// TIA Portal project "CanvasE2E" (V19)

(* hardware
DEVICE "PLC_1"  S7-1500 station
   slot 0: "导轨_0"  Rack  6ES7 590-1***0-0AA0
   slot 1: "PLC_1"  CPU 1511-1 PN  6ES7 511-1AK01-0AB0  V2.5
      slot 3: "CPU 显示_1"  6ES7591-1AA00-0AA0
      slot 32768: "PROFINET 接口_1"  X1
         slot 32769: "端口_1"  X1 P1
         slot 32770: "端口_2"  X1 P2
*)

// ===== PLC "PLC_1"  CPU 1511-1 PN =====

DATA_BLOCK "iFB_CM_CLAMP_CYL_DRV"   // DB1
{ S7_Optimized_Access := 'TRUE' }
VERSION : 0.1
// stored: InstanceOfName FB_CM_CLAMP_CYL_DRV
"FB_CM_CLAMP_CYL_DRV"
BEGIN
END_DATA_BLOCK

DATA_BLOCK "iFB_EM_CLAMP_SEQ"   // DB2
{ S7_Optimized_Access := 'TRUE' }
VERSION : 0.1
// stored: InstanceOfName FB_EM_CLAMP_SEQ
"FB_EM_CLAMP_SEQ"
BEGIN
END_DATA_BLOCK

DATA_BLOCK "iFB_U_ASSEMBLY_UNIT"   // DB3
{ S7_Optimized_Access := 'TRUE' }
VERSION : 0.1
// stored: InstanceOfName FB_U_ASSEMBLY_UNIT
"FB_U_ASSEMBLY_UNIT"
BEGIN
END_DATA_BLOCK

FUNCTION_BLOCK "PumpCtrl"   // FB1, SCL
{ S7_Optimized_Access := 'TRUE' }
   VAR_INPUT
      Start : Bool;
   END_VAR
   VAR_OUTPUT
      RunOut : Bool;
   END_VAR
   VAR
      Running : Bool;
   END_VAR
BEGIN
       // Network 1: Self-holding logic
       IF #Start THEN
           #Running := TRUE;
       END_IF;
       #RunOut := #Running;
END_FUNCTION_BLOCK

FUNCTION_BLOCK "FB_CM_CLAMP_CYL_DRV"   // FB2, SCL
{ S7_Optimized_Access := 'TRUE' }
   VAR_INPUT
      CmdExtend : Bool;
      CmdRetract : Bool;
      Extended : Bool;
      Retracted : Bool;
   END_VAR
   VAR_OUTPUT
      Q_Extend : Bool;
      Q_Retract : Bool;
      Busy : Bool;
      Done : Bool;
      Error : Bool;
   END_VAR
BEGIN
       // single-writer arbitration + feedback exclusivity
       IF #Extended AND #Retracted THEN
           #Error := TRUE;
           #Q_Extend := FALSE;
           #Q_Retract := FALSE;
       ELSE
           #Error := FALSE;
           #Q_Extend := #CmdExtend AND NOT #CmdRetract;
           #Q_Retract := #CmdRetract AND NOT #CmdExtend;
       END_IF;
       #Busy := #Q_Extend OR #Q_Retract;
END_FUNCTION_BLOCK

FUNCTION_BLOCK "FB_EM_CLAMP_SEQ"   // FB3, SCL
{ S7_Optimized_Access := 'TRUE' }
   VAR_INPUT
      Start : Bool;
      Reset : Bool;
      SafetyPermit : Bool;
      Extended : Bool;
      Retracted : Bool;
   END_VAR
   VAR_OUTPUT
      Busy : Bool;
      Done : Bool;
      Error : Bool;
      StepNo : Int;
      Extend : Bool;
      Retract : Bool;
   END_VAR
   VAR
      "Step" : Int := 0;
      FaultLatch : Bool;
      TON_S_EXTEND : TON_TIME;
      TON_S_HOLD : TON_TIME;
      TON_S_RETRACT : TON_TIME;
   END_VAR
BEGIN
       CASE #Step OF
           0: // S_WAIT 绛夊緟鍚姩
               #Busy := FALSE;
               #Done := FALSE;
               IF #Start AND #SafetyPermit THEN
                   #Step := 10;
               END_IF;
           10: // S_EXTEND 浼稿嚭澶圭揣
               #Busy := TRUE;
               #Extend := TRUE;
               #TON_S_EXTEND(IN := NOT #Extended,
                             PT := T#3000ms);
               IF #Extended THEN
                   #Extend := FALSE;
                   #Step := 20;
               END_IF;
               IF #TON_S_EXTEND.Q THEN
                   #Extend := FALSE;
                   #FaultLatch := TRUE;
                   #Step := 90;
               END_IF;
           20: // S_HOLD 淇濇寔澶圭揣
               #Busy := TRUE;
               #TON_S_HOLD(IN := TRUE,
                           PT := T#2000ms);
               IF #TON_S_HOLD.Q THEN
                   #Step := 30;
               END_IF;
           30: // S_RETRACT 缂╁洖閲婃斁
               #Busy := TRUE;
               #Retract := TRUE;
               #TON_S_RETRACT(IN := NOT #Retracted,
                              PT := T#3000ms);
               IF #Retracted THEN
                   #Retract := FALSE;
                   #Step := 40;
               END_IF;
               IF #TON_S_RETRACT.Q THEN
                   #Retract := FALSE;
                   #FaultLatch := TRUE;
                   #Step := 90;
               END_IF;
           40: // S_DONE 瀹屾垚
               #Busy := TRUE;
               #Done := TRUE;
               #Step := 0;
           90: // S_FAULT 鏁呴殰淇濇寔
               #Busy := FALSE;
               #Error := TRUE;
               #FaultLatch := TRUE;
               #Extend := FALSE;
               #Retract := FALSE;
               IF #Reset AND #Retracted AND NOT #Extended THEN
                   #FaultLatch := FALSE;
                   #Error := FALSE;
                   #Step := 0;
               END_IF;
       END_CASE;
       #StepNo := #Step;
END_FUNCTION_BLOCK

FUNCTION_BLOCK "FB_U_ASSEMBLY_UNIT"   // FB4, SCL
{ S7_Optimized_Access := 'TRUE' }
   VAR_INPUT
      Mode : Int;
      Permit : Bool;
   END_VAR
   VAR_OUTPUT
      State : Int;
      FaultSummary : Bool;
   END_VAR
BEGIN
       // shell aggregation: EM faults surface via FB_EM_*.Error (see OB_Main)
       #State := #Mode;
       #FaultSummary := FALSE;
END_FUNCTION_BLOCK

ORGANIZATION_BLOCK "Main"   // OB1, LAD, ProgramCycle
TITLE = "Main Program Sweep (Cycle)" / processos clamp cycle (LAD call shell)
{ S7_Optimized_Access := 'TRUE' }
VERSION : 0.1
   VAR_INPUT
      Initial_Call : Bool;   // Initial call of this OB
      Remanence : Bool;   // =True, if remanent data are available
   END_VAR
BEGIN

REGION Network 1
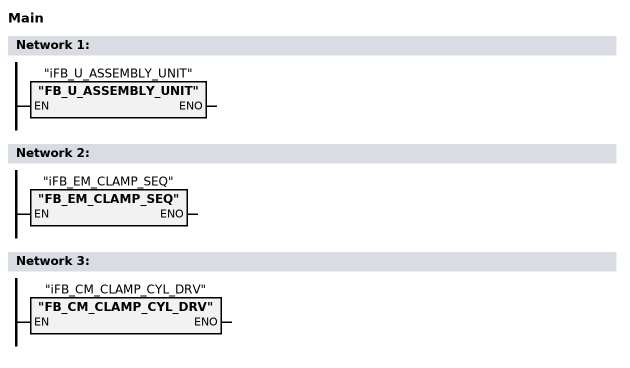
   RUNG wire#powerrail
      "iFB_U_ASSEMBLY_UNIT"()
   END_RUNG
   // the same network as SCL:
   "iFB_U_ASSEMBLY_UNIT"();   // "FB_U_ASSEMBLY_UNIT"
END_REGION

REGION Network 2
   RUNG wire#powerrail
      "iFB_EM_CLAMP_SEQ"()
   END_RUNG
   // the same network as SCL:
   "iFB_EM_CLAMP_SEQ"();   // "FB_EM_CLAMP_SEQ"
END_REGION

REGION Network 3
   RUNG wire#powerrail
      "iFB_CM_CLAMP_CYL_DRV"()
   END_RUNG
   // the same network as SCL:
   "iFB_CM_CLAMP_CYL_DRV"();   // "FB_CM_CLAMP_CYL_DRV"
END_REGION
END_ORGANIZATION_BLOCK